(* IEC 61131-3 sources: rusty/tests/lit/cfc/blocks/function_inout, 2 files *)

(* ---- addInto.st ---- *)
FUNCTION addInto : DINT
    VAR_INPUT
        delta : DINT;
    END_VAR
    VAR_IN_OUT
        acc : DINT;
    END_VAR
    acc := acc + delta;
    addInto := acc;
END_FUNCTION

(* ---- main.st ---- *)
FUNCTION main : DINT
    function_inout();
    function_inout();
    // CHECK: total = 10, result = 10
    printf('total = %d, result = %d$N', function_inout.total, function_inout.result);
END_FUNCTION
